// TIA Portal V20 export
Screen "ProductionCountSummary"  1276x673
  ScreenItem "Casella di testo_26" at 4,6 size 1273x53  Type=HmiTextBox
  ScreenItem "Casella di testo_47" at 0,0 size 881x49  Type=HmiTextBox
  ScreenItem "Casella di testo_20" at 0,50 size 97x99  Type=HmiTextBox
  ScreenItem "IO 域_1" at 99,151 size 97x49  Type=HmiIOField
  ScreenItem "IO 域_2" at 197,151 size 97x49  Type=HmiIOField
  ScreenItem "Casella di testo_8" at 0,151 size 97x49  Type=HmiTextBox
  ScreenItem "IO 域_3" at 295,151 size 97x49  Type=HmiIOField
  ScreenItem "IO 域_46" at 392,151 size 97x49  Type=HmiIOField
  ScreenItem "IO 域_47" at 491,151 size 97x49  Type=HmiIOField
  ScreenItem "IO 域_50" at 588,151 size 97x49  Type=HmiIOField
  ScreenItem "IO 域_51" at 99,201 size 97x49  Type=HmiIOField
  ScreenItem "IO 域_52" at 198,201 size 97x49  Type=HmiIOField
  ScreenItem "Casella di testo_13" at 1,201 size 97x49  Type=HmiTextBox
  ScreenItem "IO 域_55" at 296,201 size 97x49  Type=HmiIOField
  ScreenItem "IO 域_56" at 393,201 size 97x49  Type=HmiIOField
  ScreenItem "IO 域_57" at 491,201 size 97x49  Type=HmiIOField
  ScreenItem "IO 域_60" at 588,201 size 97x49  Type=HmiIOField
  ScreenItem "Casella di testo_14" at 99,101 size 97x49  Type=HmiTextBox
  ScreenItem "Casella di testo_15" at 196,101 size 97x49  Type=HmiTextBox
  ScreenItem "Casella di testo_16" at 392,101 size 97x49  Type=HmiTextBox
  ScreenItem "Casella di testo_17" at 491,101 size 97x49  Type=HmiTextBox
  ScreenItem "Casella di testo_18" at 588,101 size 97x49  Type=HmiTextBox
  ScreenItem "Casella di testo_19" at 295,101 size 97x49  Type=HmiTextBox
  ScreenItem "Casella di testo_21" at 99,50 size 194x49  Type=HmiTextBox
  ScreenItem "Casella di testo_22" at 295,50 size 194x49  Type=HmiTextBox
  ScreenItem "Casella di testo_7" at 491,50 size 389x49  Type=HmiTextBox
  ScreenItem "IO 域_61" at 99,251 size 97x49  Type=HmiIOField
  ScreenItem "IO 域_62" at 198,251 size 97x49  Type=HmiIOField
  ScreenItem "Casella di testo_23" at 1,251 size 97x49  Type=HmiTextBox
  ScreenItem "IO 域_65" at 296,251 size 97x49  Type=HmiIOField
  ScreenItem "IO 域_67" at 393,251 size 97x49  Type=HmiIOField
  ScreenItem "IO 域_70" at 491,251 size 97x49  Type=HmiIOField
  ScreenItem "IO 域_73" at 588,251 size 97x49  Type=HmiIOField
  ScreenItem "Casella di testo_1" at 686,101 size 97x49  Type=HmiTextBox
  ScreenItem "Casella di testo_2" at 783,101 size 97x49  Type=HmiTextBox
  ScreenItem "IO 域_4" at 687,151 size 97x49  Type=HmiIOField
  ScreenItem "IO 域_5" at 783,151 size 97x49  Type=HmiIOField
  ScreenItem "IO 域_6" at 687,201 size 97x49  Type=HmiIOField
  ScreenItem "IO 域_7" at 783,201 size 97x49  Type=HmiIOField
  ScreenItem "IO 域_8" at 687,251 size 97x49  Type=HmiIOField
  ScreenItem "IO 域_9" at 783,251 size 97x49  Type=HmiIOField
  ScreenItem "Casella di testo_3" at 0,0 size 881x49  Type=HmiTextBox
  ScreenItem "Casella di testo_28" at 0,51 size 97x99  Type=HmiTextBox
  ScreenItem "IO 域_20" at 99,152 size 97x49  Type=HmiIOField
  ScreenItem "IO 域_21" at 197,152 size 97x49  Type=HmiIOField
  ScreenItem "Casella di testo_29" at 0,152 size 97x49  Type=HmiTextBox
  ScreenItem "IO 域_22" at 295,152 size 97x49  Type=HmiIOField
  ScreenItem "IO 域_23" at 392,152 size 97x49  Type=HmiIOField
  ScreenItem "IO 域_24" at 491,152 size 97x49  Type=HmiIOField
  ScreenItem "IO 域_25" at 588,152 size 97x49  Type=HmiIOField
  ScreenItem "IO 域_26" at 99,202 size 97x49  Type=HmiIOField
  ScreenItem "IO 域_27" at 198,202 size 97x49  Type=HmiIOField
  ScreenItem "Casella di testo_30" at 1,202 size 97x49  Type=HmiTextBox
  ScreenItem "IO 域_28" at 296,202 size 97x49  Type=HmiIOField
  ScreenItem "IO 域_29" at 393,202 size 97x49  Type=HmiIOField
  ScreenItem "IO 域_30" at 492,202 size 97x49  Type=HmiIOField
  ScreenItem "IO 域_31" at 589,202 size 97x49  Type=HmiIOField
  ScreenItem "Casella di testo_31" at 99,102 size 97x49  Type=HmiTextBox
  ScreenItem "Casella di testo_32" at 196,102 size 97x49  Type=HmiTextBox
  ScreenItem "Casella di testo_27" at 392,102 size 97x49  Type=HmiTextBox
  ScreenItem "Casella di testo_25" at 491,102 size 97x49  Type=HmiTextBox
  ScreenItem "Casella di testo_24" at 588,102 size 97x49  Type=HmiTextBox
  ScreenItem "Casella di testo_10" at 295,102 size 97x49  Type=HmiTextBox
  ScreenItem "Casella di testo_4" at 99,51 size 194x49  Type=HmiTextBox
  ScreenItem "Casella di testo_5" at 295,51 size 194x49  Type=HmiTextBox
  ScreenItem "Casella di testo_6" at 491,51 size 389x49  Type=HmiTextBox
  ScreenItem "IO 域_10" at 99,252 size 97x49  Type=HmiIOField
  ScreenItem "IO 域_11" at 198,252 size 97x49  Type=HmiIOField
  ScreenItem "Casella di testo_9" at 1,252 size 97x49  Type=HmiTextBox
  ScreenItem "IO 域_12" at 296,252 size 97x49  Type=HmiIOField
  ScreenItem "IO 域_13" at 393,252 size 97x49  Type=HmiIOField
  ScreenItem "IO 域_19" at 492,252 size 97x49  Type=HmiIOField
  ScreenItem "IO 域_14" at 589,252 size 97x49  Type=HmiIOField
  ScreenItem "Casella di testo_11" at 686,102 size 97x49  Type=HmiTextBox
  ScreenItem "Casella di testo_12" at 783,102 size 97x49  Type=HmiTextBox
  ScreenItem "IO 域_15" at 686,152 size 97x49  Type=HmiIOField
  ScreenItem "IO 域_16" at 783,152 size 97x49  Type=HmiIOField
  ScreenItem "IO 域_17" at 687,202 size 97x49  Type=HmiIOField
  ScreenItem "IO 域_18" at 784,202 size 97x49  Type=HmiIOField
  ScreenItem "IO 域_32" at 687,252 size 97x49  Type=HmiIOField
  ScreenItem "IO 域_33" at 784,252 size 97x49  Type=HmiIOField
